(* CODESYS project iscanner.library
   Company: KOSTAL GmbH & Co.KG
   Version: 1.0.0.0
   DefaultNamespace: KOSTAL.AF2024.Drivers.Scanner.IScanner
   Title: KOSTAL.AF2024.Drivers.Scanner.IScanner
   Placeholder: KOSTAL.AF2024.Drivers.Scanner.IScanner
   Author: Frank Dümpelmann
   DocFormat: reStructuredText

Project tree, tasks and I/O mapping:
  libraries: KOSTAL.AF2024.Core.Process, 1.0.0.0 (KOSTAL GmbH & Co.KG); KOSTAL.AF2024.Core.Settings, 1.0.0.0 (KOSTAL GmbH & Co.KG); KOSTAL.AF2024.Core.System, 1.0.0.0 (KOSTAL GmbH & Co.KG)
  Interface/
    interface I_Scanner: ClearCodes, CodeGet, Ex_Scan, NativeStringGet, NumberOfBarcodes, State
  Project Information/
    function F_GetCompany [ST]
    function F_GetTitle [ST]
    function F_GetVersion [ST]
  Version/
    global variables Global_Version
*)

// Version/Global_Version
{attribute 'TcGenerated'}
{attribute 'no-analysis'}
{attribute 'linkalways'}
// This function has been automatically generated from the project information.
VAR_GLOBAL CONSTANT
	{attribute 'const_non_replaced'}
	stLibVersion_KOSTAL_AF2024_Drivers_Scanner_IScanner : ST_LibVersion := (iMajor := 1, iMinor := 0, iBuild := 0, iRevision := 0, nFlags := 0, sVersion := '1.0.0.0');
END_VAR

// Interface/I_Scanner
INTERFACE I_Scanner EXTENDS KOSTAL_AF2024_Core_System.I_Interface

METHOD ClearCodes
END_METHOD

METHOD CodeGet : KOSTAL_AF2024_Core_Settings.T_MaxString_UTF8
VAR_INPUT
	number	: UINT;
END_VAR
END_METHOD

METHOD Ex_Scan : BOOL;
VAR_INPUT
END_VAR
END_METHOD

METHOD NativeStringGet : KOSTAL_AF2024_Core_Settings.T_MaxString_UTF8
VAR_INPUT
END_VAR
END_METHOD

PROPERTY NumberOfBarcodes : UDINT
GET
END_GET
END_PROPERTY

PROPERTY State : KOSTAL_AF2024_Core_Process.I_T_PlcState
GET
END_GET
END_PROPERTY

END_INTERFACE

// Project Information/F_GetCompany
// This function has been automatically generated from the project information.
{attribute 'signature_flag' := '1073741824'}
{attribute 'TcGenerated'}
{attribute 'no-analysis'}
FUNCTION F_GetCompany : WSTRING
VAR_INPUT
	
END_VAR

F_GetCompany := "KOSTAL GmbH & Co.KG";

END_FUNCTION

// Project Information/F_GetTitle
// This function has been automatically generated from the project information.
{attribute 'signature_flag' := '1073741824'}
{attribute 'TcGenerated'}
{attribute 'no-analysis'}
FUNCTION F_GetTitle : WSTRING
VAR_INPUT
	
END_VAR

F_GetTitle := "KOSTAL.AF2024.Drivers.Scanner.IScanner";

END_FUNCTION

// Project Information/F_GetVersion
// This function has been automatically generated from the project information.
{attribute 'signature_flag' := '1073741824'}
{attribute 'TcGenerated'}
{attribute 'no-analysis'}
FUNCTION F_GetVersion : ST_LibVersion
VAR_INPUT
	
END_VAR

F_GetVersion.iMajor := 1;
F_GetVersion.iMinor := 0;
F_GetVersion.iBuild := 0;
F_GetVersion.iRevision := 0;
F_GetVersion.sVersion := '1.0.0.0';
F_GetVersion.nFlags := 0;

END_FUNCTION
